TYPE ST_ExampleStationConfiguration :
STRUCT
	cycleDwell			: TIME := T#2S; //wait time between jobs while running
	maxCloseDwell		: TIME := T#10S; //longest closeDwell accepted in a request
END_STRUCT
END_TYPE

(* stored: Version 1.1.0.1, ProductVersion 3.1.4024.12
   DUT ST_ExampleStationConfiguration: Id {434ce971-85e6-4397-9a11-c884bb9f974f} *)
